Fanuc KAREL source: KC00014.KL

PROGRAM KC00014
%NOLOCKGROUP
%ENVIRONMENT TIM
VAR
  I: INTEGER
  J: INTEGER
  K: INTEGER
  R: REAL
  B: BOOLEAN
  S: STRING[80]
  T: STRING[80]
  P: PATH
  Q: PATH
  AI: ARRAY[8] OF INTEGER
  AB: ARRAY[244] OF BYTE
BEGIN
  I = GET_USEC_TIM
END KC00014
